(* IEC 61131-3 sources: SRCI_CLIENT_PLC/RobotLibrary/Library/Structures/Axis, 4 files *)

(* ---- AxisExternalUnit.st ---- *)
TYPE AxisExternalUnit :
// -------------------------------------------------------------------------
//  SRCI Robot Library
// -------------------------------------------------------------------------
//
//  Object:      AxisExternalUnit
//  Author:      Thorsten Brach
//  Date:        2025-03-23
//
//  Description:
//
//
//  Copyright:
//    (C) 2025 Thorsten Brach. All rights reserved
//             Licensed under the MIT License.
//
//  Disclaimer:
//    This project is provided without any guarantee and can be used for
//    private and commercial purposes. Any use is at the user’s
//    own risk and responsibility.
//
// -------------------------------------------------------------------------
STRUCT
  /// External Axis 1 used
  E1 : AxisUnit;
  /// External Axis 2 used
  E2 : AxisUnit;
  /// External Axis 3 used
  E3 : AxisUnit;
  /// External Axis 4 used
  E4 : AxisUnit;
  /// External Axis 5 used
  E5 : AxisUnit;
  /// External Axis 6 used
  E6 : AxisUnit;
END_STRUCT
END_TYPE

(* ---- AxisExternalUsed.st ---- *)
TYPE AxisExternalUsed :
// -------------------------------------------------------------------------
//  SRCI Robot Library
// -------------------------------------------------------------------------
//
//  Object:      AxisExternalUsed
//  Author:      Thorsten Brach
//  Date:        2025-03-23
//
//  Description:
//
//
//  Copyright:
//    (C) 2025 Thorsten Brach. All rights reserved
//             Licensed under the MIT License.
//
//  Disclaimer:
//    This project is provided without any guarantee and can be used for
//    private and commercial purposes. Any use is at the user’s
//    own risk and responsibility.
//
// -------------------------------------------------------------------------
STRUCT
  /// External Axis 1 used
  E1 : BOOL;
  /// External Axis 2 used
  E2 : BOOL;
  /// External Axis 3 used
  E3 : BOOL;
  /// External Axis 4 used
  E4 : BOOL;
  /// External Axis 5 used
  E5 : BOOL;
  /// External Axis 6 used
  E6 : BOOL;
END_STRUCT
END_TYPE

(* ---- AxisJointUnit.st ---- *)
TYPE AxisJointUnit :
// -------------------------------------------------------------------------
//  SRCI Robot Library
// -------------------------------------------------------------------------
//
//  Object:      AxisJointUnit
//  Author:      Thorsten Brach
//  Date:        2025-03-23
//
//  Description:
//
//
//  Copyright:
//    (C) 2025 Thorsten Brach. All rights reserved
//             Licensed under the MIT License.
//
//  Disclaimer:
//    This project is provided without any guarantee and can be used for
//    private and commercial purposes. Any use is at the user’s
//    own risk and responsibility.
//
// -------------------------------------------------------------------------
STRUCT
  /// Joint Axis 1 unit
  J1 : AxisUnit;
  /// Joint Axis 2 unit
  J2 : AxisUnit;
  /// Joint Axis 3 unit
  J3 : AxisUnit;
  /// Joint Axis 4 unit
  J4 : AxisUnit;
  /// Joint Axis 5 unit
  J5 : AxisUnit;
  /// Joint Axis 6 unit
  J6 : AxisUnit;
END_STRUCT
END_TYPE

(* ---- AxisJointUsed.st ---- *)
TYPE AxisJointUsed :
// -------------------------------------------------------------------------
//  SRCI Robot Library
// -------------------------------------------------------------------------
//
//  Object:      AxisJointUsed
//  Author:      Thorsten Brach
//  Date:        2025-03-23
//
//  Description:
//
//
//  Copyright:
//    (C) 2025 Thorsten Brach. All rights reserved
//             Licensed under the MIT License.
//
//  Disclaimer:
//    This project is provided without any guarantee and can be used for
//    private and commercial purposes. Any use is at the user’s
//    own risk and responsibility.
//
// -------------------------------------------------------------------------
STRUCT
  /// Joint Axis 1 used
  J1 : BOOL;
  /// Joint Axis 2 used
  J2 : BOOL;
  /// Joint Axis 3 used
  J3 : BOOL;
  /// Joint Axis 4 used
  J4 : BOOL;
  /// Joint Axis 5 used
  J5 : BOOL;
  /// Joint Axis 6 used
  J6 : BOOL;
END_STRUCT
END_TYPE
